RoboDK station: cell_station.rdk

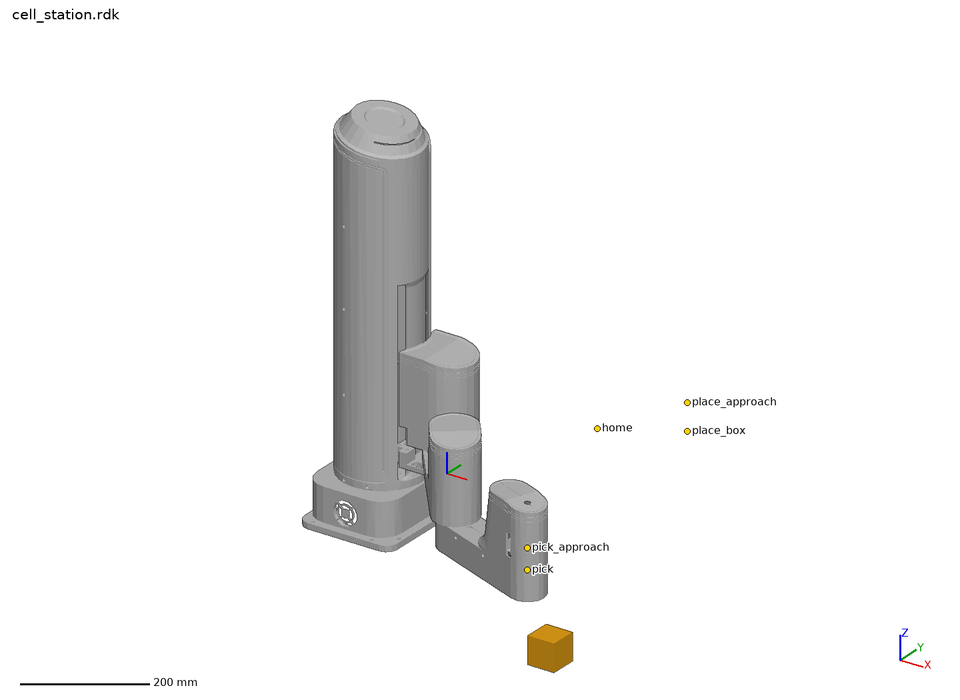
[picture v0: the station drawn from its stored meshes, robots at their saved joint values, targets as dots, program paths as lines]
Station cell_station (saved by RoboDK 5.9.6). Poses are relative to the parent item; angles as X-Y-Z fixed-axis rotations.
  - frame Dobot M1 Base at (0, 0, 0) mm
    - robot Dobot M1: 4 axes, payload 1.5 kg, reach 446 mm, repeatability 0.01 mm, weight 14 kg
        modified DH rows (alpha deg, a mm, theta deg, d mm): 0, 0, 0, -53 linear; 0, 0, 0, 0; 0, 200, 0, 0; 180, 200, 0, 0
        joint limits [0, -90, -135, -180] to [250, 90, 135, 180]; home [200, -45, 90, 45]; saved at [15.73, -51.34, 30.11, 7.77]
      - tool vacuum cup, TCP at (0, 0, -50) mm
    - target home (Cartesian target) at (282.84, 0, 157) mm, rotated rx 180 ry 0 rz 0 deg; joints [160, -45, 90, 45] of Dobot M1
    - target pick (Cartesian target) at (311.37, -228.6, 12.73) mm, rotated rx 180 ry 0 rz -29 deg; joints [15.73, -51.34, 30.11, 7.77] of Dobot M1
    - target pick_approach (Cartesian target) at (311.37, -228.6, 50.73) mm, rotated rx 180 ry 0 rz -29 deg; joints [53.73, -51.34, 30.11, 7.77] of Dobot M1
    - target place_box (Cartesian target) at (305.83, 210.47, 73.92) mm, rotated rx 180 ry 0 rz 56.39 deg; joints [76.92, 12.68, 43.71, 0] of Dobot M1
    - target place_approach (Cartesian target) at (305.83, 210.47, 123.92) mm, rotated rx 180 ry 0 rz 56.39 deg; joints [126.92, 12.68, 43.71, 0] of Dobot M1
  - object item at (311, -228, -150) mm, size 50 x 50 x 50 mm, geometry from Cube-50mm.sld
